{attribute 'qualified_only'}
{attribute 'strict'}
{attribute 'to_string'}
TYPE E_FillStep :
(
    Undefined := 0,
    Idle      := 10,
    Opening   := 20,
    Filling   := 30,
    Closing   := 40,
    Done      := 50,
    Error     := 900
);
END_TYPE

(* stored: Version 1.1.0.1
   DUT E_FillStep: Id {1fd7d39b-76d7-48c7-bb74-e46758d835c3} *)
